FUNCTION_BLOCK FB_ConveyorTracking4Pt
VAR_INPUT
    bResetSystem     : BOOL;
    bCameraResult    : BOOL;
    rCenterX_mm      : LREAL;
    rCenterY_mm      : LREAL;
    rAngleDeg        : LREAL;
    rLength_mm       : LREAL := 40.0;
    rWidth_mm        : LREAL := 40.0;
    nEncoderNow      : UINT;
    rMmPerPulse      : LREAL := 0.476475;
    rXMaxLimit_mm    : LREAL := 180.0;
END_VAR

VAR_OUTPUT
    bProductValid    : BOOL;
    nPulseAtCamera   : UINT;
    nPulseTravel     : INT;
    rTravel_mm       : LREAL;
    aCornerBase      : ARRAY[1..4] OF ST_Point2D;
    aCornerNow       : ARRAY[1..4] OF ST_Point2D;
END_VAR

VAR
    fbCameraEdge     : R_TRIG;
    rRad             : LREAL;
    rCosA            : LREAL;
    rSinA            : LREAL;
    rHalfLength      : LREAL;
    rHalfWidth       : LREAL;
    nIndex           : INT;
    bFirstScan       : BOOL := TRUE;
END_VAR

// Reset mốc phần mềm một lần khi PLC khởi động hoặc khi bResetSystem kích.
IF bFirstScan OR bResetSystem THEN
    bFirstScan     := FALSE;
    bProductValid  := FALSE;
    nPulseAtCamera := nEncoderNow;
    nPulseTravel   := 0;
    rTravel_mm     := 0.0;

    FOR nIndex := 1 TO 4 DO
        aCornerBase[nIndex].X := 0.0;
        aCornerBase[nIndex].Y := 0.0;
        aCornerNow[nIndex].X  := 0.0;
        aCornerNow[nIndex].Y  := 0.0;
    END_FOR;
END_IF;

fbCameraEdge(CLK := bCameraResult);

// Camera chụp: chốt encoder và tính bốn góc gốc.
IF fbCameraEdge.Q THEN
    nPulseAtCamera := nEncoderNow;
    nPulseTravel   := 0;
    rTravel_mm     := 0.0;

    rRad   := rAngleDeg * 3.141592653589793 / 180.0;
    rCosA  := COS(rRad);
    rSinA  := SIN(rRad);
    rHalfLength := rLength_mm / 2.0;
    rHalfWidth  := rWidth_mm / 2.0;

    aCornerBase[1].X := rCenterX_mm + rHalfLength * rCosA - rHalfWidth * rSinA;
    aCornerBase[1].Y := rCenterY_mm + rHalfLength * rSinA + rHalfWidth * rCosA;
    aCornerBase[2].X := rCenterX_mm - rHalfLength * rCosA - rHalfWidth * rSinA;
    aCornerBase[2].Y := rCenterY_mm - rHalfLength * rSinA + rHalfWidth * rCosA;
    aCornerBase[3].X := rCenterX_mm - rHalfLength * rCosA + rHalfWidth * rSinA;
    aCornerBase[3].Y := rCenterY_mm - rHalfLength * rSinA - rHalfWidth * rCosA;
    aCornerBase[4].X := rCenterX_mm + rHalfLength * rCosA + rHalfWidth * rSinA;
    aCornerBase[4].Y := rCenterY_mm + rHalfLength * rSinA - rHalfWidth * rCosA;

    FOR nIndex := 1 TO 4 DO
        aCornerNow[nIndex] := aCornerBase[nIndex];
    END_FOR;
    bProductValid := TRUE;
END_IF;

// Tracking thời gian thực theo encoder.
IF bProductValid THEN
    nPulseTravel := TO_INT(nEncoderNow - nPulseAtCamera);
    rTravel_mm   := TO_LREAL(nPulseTravel) * rMmPerPulse;

    FOR nIndex := 1 TO 4 DO
        aCornerNow[nIndex].X := aCornerBase[nIndex].X + rTravel_mm;
        aCornerNow[nIndex].Y := aCornerBase[nIndex].Y;
    END_FOR;

    // Hủy sản phẩm nếu toàn bộ cạnh phía sau đã vượt vùng X của Gantry.
    IF (aCornerNow[2].X > rXMaxLimit_mm) AND (aCornerNow[3].X > rXMaxLimit_mm) THEN
        bProductValid := FALSE;
        nPulseTravel  := 0;
        rTravel_mm    := 0.0;
    END_IF;
END_IF;

END_FUNCTION_BLOCK

(* stored: Version 1.1.0.1, ProductVersion 3.1.4024.16
   POU FB_ConveyorTracking4Pt: Id {f45dd975-916c-42e3-9485-f5e77a4a0ab5}, SpecialFunc None *)
